// TIA Portal V20 export
// export: Created 2026-10-12T16:46:21.1158683Z, ExportSetting WithDefaults, DisplayName Totally Integrated Automation Portal, DisplayVersion V20 Update 6, DisplayName TIA Portal Openness, DisplayVersion V20 Update 6, DisplayName TIA Portal Version Control Interface, DisplayVersion V20 Update 6, DisplayName SINAMICS Startdrive Advanced, DisplayVersion V20 SP1 Update 2, DisplayName SINAMICS Startdrive G110M, G120, G120C, G120D, G120P, G115D, DisplayVersion V20 SP1 Update 2, DisplayName SINAMICS Startdrive G130, G150, S120, S150, SINAMICS MV, G220, S200, S210, DisplayVersion V20 SP1 Update 2, DisplayName STEP 7 Professional, DisplayVersion V20 Update 6, DisplayName STEP 7 Safety, DisplayVersion V20 Update 2, DisplayName WinCC Basic/Comfort/Advanced, DisplayVersion V20 Update 6, DisplayName WinCC Professional, DisplayVersion V20 Update 6, DisplayName WinCC Unified, DisplayVersion V20 Update 6
DATA_BLOCK "DB_Fehlermeldungen"   // DB39
{ S7_Optimized_Access := 'TRUE' }
VERSION : 0.2
// FI-Schutz ausgeloest (Heizungen)
// stored: AutoNumber true, DBAccessibleFromOPCUA true, DBAccessibleFromWebserver true, IsOnlyStoredInLoadMemory false, IsRetainMemResEnabled false, IsWriteProtectedInAS false, MemoryReserve 100
   VAR
      FI_Heizung_Bad_7 : Bool;   // 1 - FI-Schutz 200F1 Heizung Bad 7 ausgeloest
      FI_Heizung_Bad_8 : Bool;   // 2 - FI-Schutz 210F1 Heizung Bad 8 ausgeloest
      FI_Heizung_Bad_12 : Bool;   // 3 - FI-Schutz 220F1 Heizung Bad 12 ausgeloest
      FI_Heizung_Bad_25 : Bool;   // 4 - FI+Motorschutz 270/271 Heizung Bad 25 ausgeloest
      FI_Heizung_Bad_36 : Bool;   // 5 - FI-Schutz 300F1 Heizung Bad 36 ausgeloest
      FI_Heizung_Bad_40 : Bool;   // 6 - FI-Schutz 310F1 Heizung Bad 40 ausgeloest
      FI_Heizung_Bad_46 : Bool;   // 7 - FI-Schutz 340F1 Heizung Bad 46 ausgeloest Uebertemperatur (Heizungen)
      Uebertemp_Bad_7 : Bool;   // 8 - Uebertemperatur Heizung Bad 7
      Uebertemp_Bad_8 : Bool;   // 9 - Uebertemperatur Heizung Bad 8
      Uebertemp_Bad_12 : Bool;   // 10 - Uebertemperatur Heizung Bad 12
      Uebertemp_Bad_25 : Bool;   // 11 - Uebertemperatur Heizung Bad 25
      Uebertemp_Bad_36 : Bool;   // 12 - Uebertemperatur Heizung Bad 36
      Uebertemp_Bad_40 : Bool;   // 13 - Uebertemperatur Heizung Bad 40
      Uebertemp_Bad_46 : Bool;   // 14 - Uebertemperatur Heizung Bad 46 Motorschutz Pumpe ausgeloest
      Motorschutz_Pumpe_Bad_8 : Bool;   // 15 - Motorschutz 215Q1 Pumpe Bad 8 ausgeloest
      Motorschutz_Pumpe_Bad_12 : Bool;   // 16 - Motorschutz 225Q1 Pumpe Bad 12 ausgeloest
      Motorschutz_Pumpe_Bad_14 : Bool;   // 17 - Motorschutz 235Q1 Pumpe Bad 14 ausgeloest
      Motorschutz_Pumpe_Bad_18 : Bool;   // 18 - Motorschutz 245Q1 Pumpe Bad 18 ausgeloest
      Motorschutz_Pumpe_Bad_19 : Bool;   // 19 - Motorschutz 255Q1 Pumpe Bad 19 ausgeloest
      Motorschutz_Pumpe_Bad_21 : Bool;   // 20 - Motorschutz 265Q1 Pumpe Bad 21 ausgeloest
      Motorschutz_Pumpe_Bad_25 : Bool;   // 21 - Motorschutz 275Q1 Pumpe Bad 25 ausgeloest
      Motorschutz_Pumpe_Bad_26 : Bool;   // 22 - Motorschutz 285Q1 Pumpe Bad 26 ausgeloest
      Motorschutz_Pumpe_Bad_31 : Bool;   // 23 - Motorschutz 295Q1 Pumpe Bad 31 ausgeloest
      Motorschutz_Pumpe_Bad_41 : Bool;   // 24 - Motorschutz 325Q1 Pumpe Bad 41 ausgeloest
      Motorschutz_Pumpe_Bad_45 : Bool;   // 25 - Motorschutz 335Q1 Pumpe Bad 45 ausgeloest Wartungsschalter Pumpe nicht eingeschaltet
      Wartungsschalter_Pumpe_Bad_8 : Bool;   // 26 - Wartungsschalter Pumpe Bad 8 nicht eingeschaltet
      Wartungsschalter_Pumpe_Bad_12 : Bool;   // 27 - Wartungsschalter Pumpe Bad 12 nicht eingeschaltet
      Wartungsschalter_Pumpe_Bad_14 : Bool;   // 28 - Wartungsschalter Pumpe Bad 14 nicht eingeschaltet
      Wartungsschalter_Pumpe_Bad_18 : Bool;   // 29 - Wartungsschalter Pumpe Bad 18 nicht eingeschaltet
      Wartungsschalter_Pumpe_Bad_19 : Bool;   // 30 - Wartungsschalter Pumpe Bad 19 nicht eingeschaltet
      Wartungsschalter_Pumpe_Bad_21 : Bool;   // 31 - Wartungsschalter Pumpe Bad 21 nicht eingeschaltet
      Wartungsschalter_Pumpe_Bad_25 : Bool;   // 32 - Wartungsschalter Pumpe Bad 25 nicht eingeschaltet
      Wartungsschalter_Pumpe_Bad_26 : Bool;   // 33 - Wartungsschalter Pumpe Bad 26 nicht eingeschaltet
      Wartungsschalter_Pumpe_Bad_31 : Bool;   // 34 - Wartungsschalter Pumpe Bad 31 nicht eingeschaltet
      Wartungsschalter_Pumpe_Bad_41 : Bool;   // 35 - Wartungsschalter Pumpe Bad 41 nicht eingeschaltet
      Wartungsschalter_Pumpe_Bad_45 : Bool;   // 36 - Wartungsschalter Pumpe Bad 45 nicht eingeschaltet Niveau nicht OK
      Niveau_Bad_7 : Bool;   // 37 - Niveau Bad 7 nicht OK
      Niveau_Bad_8 : Bool;   // 38 - Niveau Bad 8 nicht OK
      Niveau_Bad_12 : Bool;   // 39 - Niveau Bad 12 nicht OK
      Niveau_Bad_25 : Bool;   // 40 - Niveau Bad 25 nicht OK
      Niveau_Bad_36 : Bool;   // 41 - Niveau Bad 36 nicht OK
      Niveau_Bad_40 : Bool;   // 42 - Niveau Bad 40 nicht OK
      Niveau_Bad_46 : Bool;   // 43 - Niveau Bad 46 nicht OK Frequenzumrichter Stoerung (angesteuert aber nicht bereit, 3s verzoegert)
      FU_Pumpe_Bad_25 : Bool;   // 44 - FU Umwaelzpumpe Bad 25 Stoerung
      FU_WB1_Bad_25 : Bool;   // 45 - FU Warenbewegung 1 Bad 25 Stoerung
      FU_WB2_Bad_25 : Bool;   // 46 - FU Warenbewegung 2 Bad 25 Stoerung Motorschutz Warenbewegung ausgeloest
      Motorschutz_WB1_Bad_25 : Bool;   // 47 - Motorschutz 276Q1 Warenbewegung 1 Bad 25 ausgeloest
      Motorschutz_WB2_Bad_25 : Bool;   // 48 - Motorschutz 277Q1 Warenbewegung 2 Bad 25 ausgeloest PT100 Sensorstoerung (Drahtbruch oder Kurzschluss)
      PT100_Bad_7 : Bool;   // 49 - PT100 Heizung Bad 7 Sensorstoerung
      PT100_Bad_8 : Bool;   // 50 - PT100 Heizung Bad 8 Sensorstoerung
      PT100_Bad_12 : Bool;   // 51 - PT100 Heizung Bad 12 Sensorstoerung
      PT100_Bad_25_H1 : Bool;   // 52 - PT100 Heizung 1 Bad 25 Sensorstoerung
      PT100_Bad_25_H2 : Bool;   // 53 - PT100 Heizung 2 Bad 25 Sensorstoerung
      PT100_Bad_36 : Bool;   // 54 - PT100 Heizung Bad 36 Sensorstoerung
      PT100_Bad_40 : Bool;   // 55 - PT100 Heizung Bad 40 Sensorstoerung
      PT100_Bad_46 : Bool;   // 56 - PT100 Heizung Bad 46 Sensorstoerung Walchem Controller
      Fehler_Walchem_Controller : Bool;   // 57 - Alarm Walchem Controller Bad 25 Not-Halt
      Not_Halt : Bool;   // 58 - Not-Halt ausgeloest
   END_VAR
BEGIN
END_DATA_BLOCK
